// TIA Portal V19 export
FUNCTION_BLOCK "ALL HOOTER"   // FB9, LAD
{ S7_Optimized_Access := 'TRUE' }
// stored: MemoryReserve 100, SetENOAutomatically false
   VAR
      HOOTER_Instance { S7_SetPoint := 'True'} : "HOOTER";
      HOOTER_Instance_1 { S7_SetPoint := 'True'} : "HOOTER";
   END_VAR
   VAR_TEMP   // added for the SCL form of the ladder/FBD networks
      _w1 : Bool;
      _w2 : Bool;
   END_VAR
BEGIN

REGION Network 1
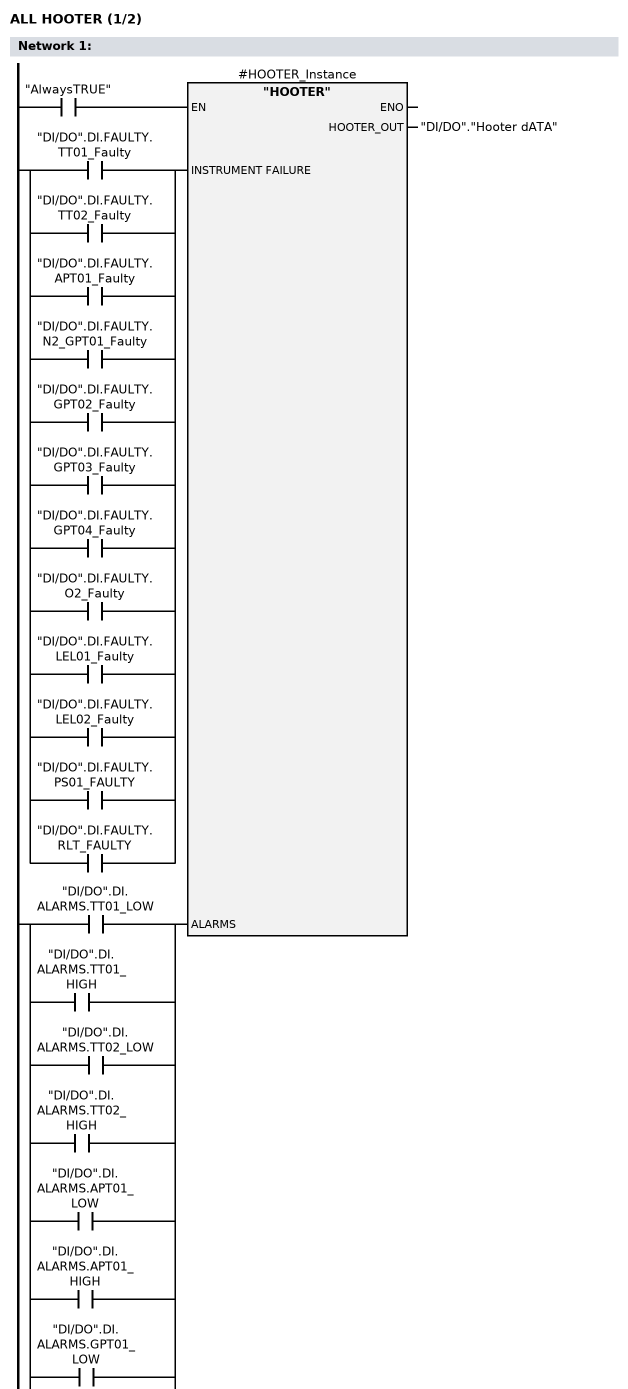
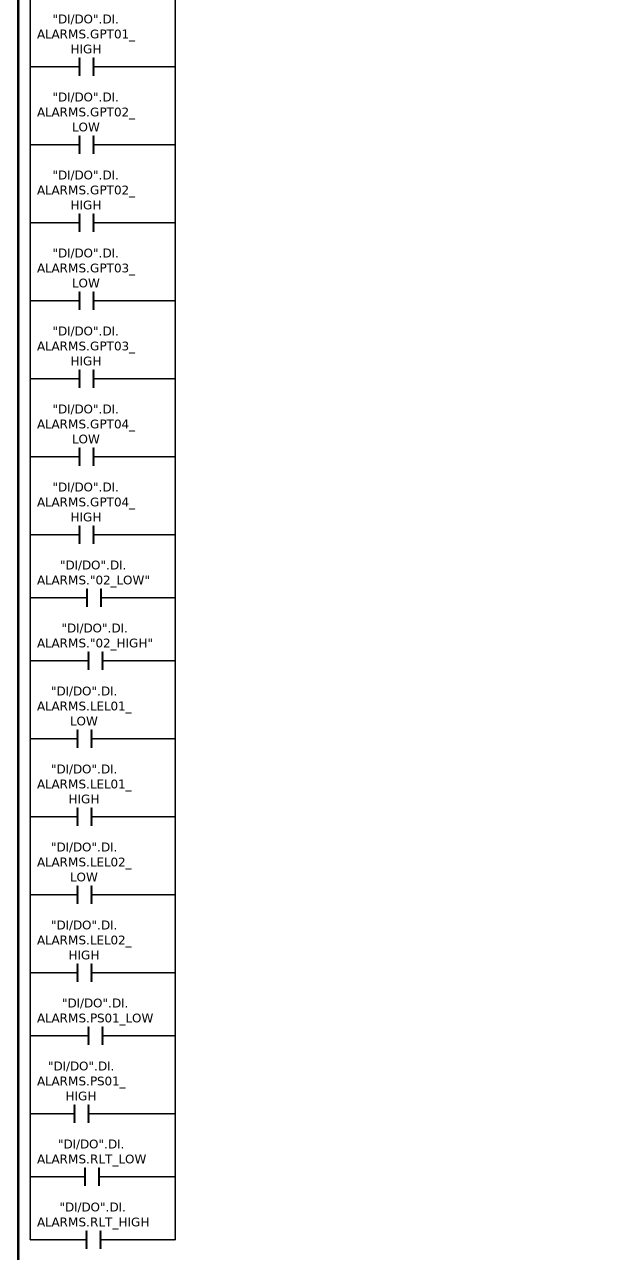
   RUNG wire#powerrail
      Contact( "AlwaysTRUE" )
      #HOOTER_Instance("INSTRUMENT FAILURE" := wire#w1, ALARMS := wire#w2, HOOTER_OUT => "DI/DO"."Hooter dATA")
   END_RUNG
   RUNG wire#powerrail
      Contact( "DI/DO".DI.FAULTY.TT01_Faulty )
   END_RUNG wire#w1
   RUNG wire#powerrail
      Contact( "DI/DO".DI.FAULTY.TT02_Faulty )
   END_RUNG wire#w1
   RUNG wire#powerrail
      Contact( "DI/DO".DI.FAULTY.APT01_Faulty )
   END_RUNG wire#w1
   RUNG wire#powerrail
      Contact( "DI/DO".DI.FAULTY.N2_GPT01_Faulty )
   END_RUNG wire#w1
   RUNG wire#powerrail
      Contact( "DI/DO".DI.FAULTY.GPT02_Faulty )
   END_RUNG wire#w1
   RUNG wire#powerrail
      Contact( "DI/DO".DI.FAULTY.GPT03_Faulty )
   END_RUNG wire#w1
   RUNG wire#powerrail
      Contact( "DI/DO".DI.FAULTY.GPT04_Faulty )
   END_RUNG wire#w1
   RUNG wire#powerrail
      Contact( "DI/DO".DI.FAULTY.O2_Faulty )
   END_RUNG wire#w1
   RUNG wire#powerrail
      Contact( "DI/DO".DI.FAULTY.LEL01_Faulty )
   END_RUNG wire#w1
   RUNG wire#powerrail
      Contact( "DI/DO".DI.FAULTY.LEL02_Faulty )
   END_RUNG wire#w1
   RUNG wire#powerrail
      Contact( "DI/DO".DI.FAULTY.PS01_FAULTY )
   END_RUNG wire#w1
   RUNG wire#powerrail
      Contact( "DI/DO".DI.FAULTY.RLT_FAULTY )
   END_RUNG wire#w1
   RUNG wire#powerrail
      Contact( "DI/DO".DI.ALARMS.TT01_LOW )
   END_RUNG wire#w2
   RUNG wire#powerrail
      Contact( "DI/DO".DI.ALARMS.TT01_HIGH )
   END_RUNG wire#w2
   RUNG wire#powerrail
      Contact( "DI/DO".DI.ALARMS.TT02_LOW )
   END_RUNG wire#w2
   RUNG wire#powerrail
      Contact( "DI/DO".DI.ALARMS.TT02_HIGH )
   END_RUNG wire#w2
   RUNG wire#powerrail
      Contact( "DI/DO".DI.ALARMS.APT01_LOW )
   END_RUNG wire#w2
   RUNG wire#powerrail
      Contact( "DI/DO".DI.ALARMS.APT01_HIGH )
   END_RUNG wire#w2
   RUNG wire#powerrail
      Contact( "DI/DO".DI.ALARMS.GPT01_LOW )
   END_RUNG wire#w2
   RUNG wire#powerrail
      Contact( "DI/DO".DI.ALARMS.GPT01_HIGH )
   END_RUNG wire#w2
   RUNG wire#powerrail
      Contact( "DI/DO".DI.ALARMS.GPT02_LOW )
   END_RUNG wire#w2
   RUNG wire#powerrail
      Contact( "DI/DO".DI.ALARMS.GPT02_HIGH )
   END_RUNG wire#w2
   RUNG wire#powerrail
      Contact( "DI/DO".DI.ALARMS.GPT03_LOW )
   END_RUNG wire#w2
   RUNG wire#powerrail
      Contact( "DI/DO".DI.ALARMS.GPT03_HIGH )
   END_RUNG wire#w2
   RUNG wire#powerrail
      Contact( "DI/DO".DI.ALARMS.GPT04_LOW )
   END_RUNG wire#w2
   RUNG wire#powerrail
      Contact( "DI/DO".DI.ALARMS.GPT04_HIGH )
   END_RUNG wire#w2
   RUNG wire#powerrail
      Contact( "DI/DO".DI.ALARMS."02_LOW" )
   END_RUNG wire#w2
   RUNG wire#powerrail
      Contact( "DI/DO".DI.ALARMS."02_HIGH" )
   END_RUNG wire#w2
   RUNG wire#powerrail
      Contact( "DI/DO".DI.ALARMS.LEL01_LOW )
   END_RUNG wire#w2
   RUNG wire#powerrail
      Contact( "DI/DO".DI.ALARMS.LEL01_HIGH )
   END_RUNG wire#w2
   RUNG wire#powerrail
      Contact( "DI/DO".DI.ALARMS.LEL02_LOW )
   END_RUNG wire#w2
   RUNG wire#powerrail
      Contact( "DI/DO".DI.ALARMS.LEL02_HIGH )
   END_RUNG wire#w2
   RUNG wire#powerrail
      Contact( "DI/DO".DI.ALARMS.PS01_LOW )
   END_RUNG wire#w2
   RUNG wire#powerrail
      Contact( "DI/DO".DI.ALARMS.PS01_HIGH )
   END_RUNG wire#w2
   RUNG wire#powerrail
      Contact( "DI/DO".DI.ALARMS.RLT_LOW )
   END_RUNG wire#w2
   RUNG wire#powerrail
      Contact( "DI/DO".DI.ALARMS.RLT_HIGH )
   END_RUNG wire#w2
   // the same network as SCL:
   IF "AlwaysTRUE" THEN
       #HOOTER_Instance("INSTRUMENT FAILURE" := "DI/DO".DI.FAULTY.TT01_Faulty OR "DI/DO".DI.FAULTY.TT02_Faulty OR "DI/DO".DI.FAULTY.APT01_Faulty OR "DI/DO".DI.FAULTY.N2_GPT01_Faulty OR "DI/DO".DI.FAULTY.GPT02_Faulty OR "DI/DO".DI.FAULTY.GPT03_Faulty OR "DI/DO".DI.FAULTY.GPT04_Faulty OR "DI/DO".DI.FAULTY.O2_Faulty OR "DI/DO".DI.FAULTY.LEL01_Faulty OR "DI/DO".DI.FAULTY.LEL02_Faulty OR "DI/DO".DI.FAULTY.PS01_FAULTY OR "DI/DO".DI.FAULTY.RLT_FAULTY,   // "HOOTER"
                        ALARMS := "DI/DO".DI.ALARMS.TT01_LOW OR "DI/DO".DI.ALARMS.TT01_HIGH OR "DI/DO".DI.ALARMS.TT02_LOW OR "DI/DO".DI.ALARMS.TT02_HIGH OR "DI/DO".DI.ALARMS.APT01_LOW OR "DI/DO".DI.ALARMS.APT01_HIGH OR "DI/DO".DI.ALARMS.GPT01_LOW OR "DI/DO".DI.ALARMS.GPT01_HIGH OR "DI/DO".DI.ALARMS.GPT02_LOW OR "DI/DO".DI.ALARMS.GPT02_HIGH OR "DI/DO".DI.ALARMS.GPT03_LOW OR "DI/DO".DI.ALARMS.GPT03_HIGH OR "DI/DO".DI.ALARMS.GPT04_LOW OR "DI/DO".DI.ALARMS.GPT04_HIGH OR "DI/DO".DI.ALARMS."02_LOW" OR "DI/DO".DI.ALARMS."02_HIGH" OR "DI/DO".DI.ALARMS.LEL01_LOW OR "DI/DO".DI.ALARMS.LEL01_HIGH OR "DI/DO".DI.ALARMS.LEL02_LOW OR "DI/DO".DI.ALARMS.LEL02_HIGH OR "DI/DO".DI.ALARMS.PS01_LOW OR "DI/DO".DI.ALARMS.PS01_HIGH OR "DI/DO".DI.ALARMS.RLT_LOW OR "DI/DO".DI.ALARMS.RLT_HIGH,
                        HOOTER_OUT => "DI/DO"."Hooter dATA");
   END_IF;
END_REGION

REGION Network 2
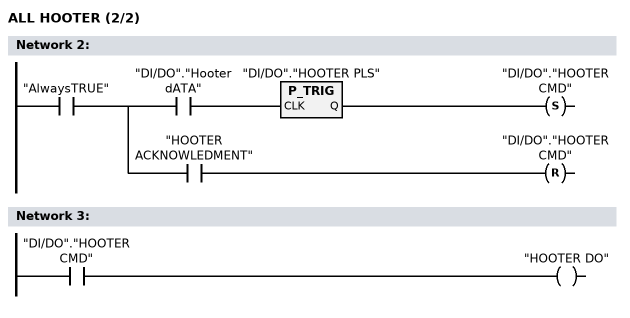
   RUNG wire#powerrail
      Contact( "AlwaysTRUE" )
      wire#w1
      Contact( "DI/DO"."Hooter dATA" )
      P_Trig( "DI/DO"."HOOTER PLS" )
      S_Coil( "DI/DO"."HOOTER CMD" )
   END_RUNG
   RUNG wire#w1
      Contact( "HOOTER ACKNOWLEDMENT" )
      R_Coil( "DI/DO"."HOOTER CMD" )
   END_RUNG
   // the same network as SCL:
   #_w1 := "AlwaysTRUE" AND "DI/DO"."Hooter dATA";
   #_w2 := #_w1 AND NOT "DI/DO"."HOOTER PLS";   // rising edge
   "DI/DO"."HOOTER PLS" := #_w1;
   IF #_w2 THEN "DI/DO"."HOOTER CMD" := TRUE; END_IF;
   IF "AlwaysTRUE" AND "HOOTER ACKNOWLEDMENT" THEN "DI/DO"."HOOTER CMD" := FALSE; END_IF;
END_REGION

REGION Network 3
   RUNG wire#powerrail
      Contact( "DI/DO"."HOOTER CMD" )
      Coil( "HOOTER DO" )
   END_RUNG
   // the same network as SCL:
   "HOOTER DO" := "DI/DO"."HOOTER CMD";
END_REGION
END_FUNCTION_BLOCK
